% RSLogix 500 project PROGRAM_-7_BAK017.RSS, saved by version 8.30.00.16 %
PROJECT "UNTITLED"    % processor: Bul.1763 MicroLogix 1100 Series B %

PROGRAM FILES
  LAD 2 "MAIN"  4 rungs
  LAD 3 "IO"  4 rungs
  LAD 4 "SAMPL_CYCL"  2 rungs
  LAD 5 "CAL_CYCL"  14 rungs

DATA FILES
  O0 OUTPUT  4 elements
  I1 INPUT  6 elements
  S2 STATUS  66 elements
  B3 BINARY  1 elements
  T4 TIMER  3 elements
  C5 COUNTER  1 elements
  R6 CONTROL  1 elements
  N7 INTEGER  8 elements
  F8 FLOAT  7 elements

LADDER 2 "MAIN"
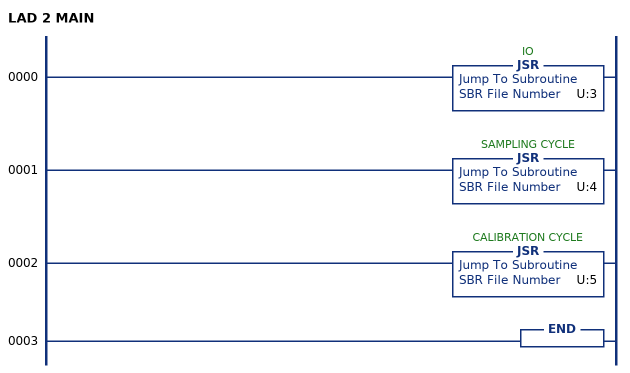
% Rung: 0 %
SOR JSR U:3 EOR
%   U:3  "IO" %
% Rung: 1 %
SOR JSR U:4 EOR
%   U:4  "SAMPLING CYCLE" %
% Rung: 2 %
SOR JSR U:5 EOR
%   U:5  "CALIBRATION CYCLE" %
% Rung: 3 %
SOR END EOR

LADDER 3 "IO"
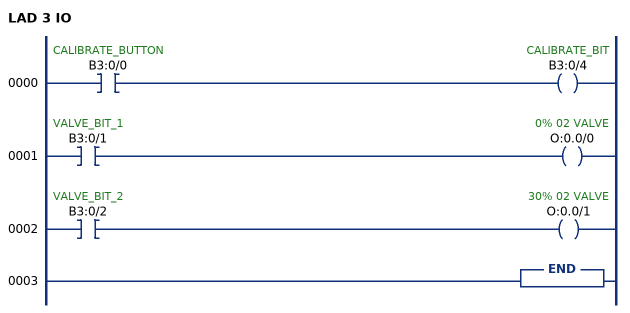
% Rung: 0 %
SOR XIC B3:0/0 OTE B3:0/4 EOR
%   B3:0/0  CALIBRATE_BUTTON %
%   B3:0/4  CALIBRATE_BIT %
% Rung: 1 %
SOR XIC B3:0/1 OTE O:0.0/0 EOR
%   B3:0/1  VALVE_BIT_1 %
%   O:0.0/0  "0% 02 VALVE" %
% Rung: 2 %
SOR XIC B3:0/2 OTE O:0.0/1 EOR
%   B3:0/2  VALVE_BIT_2 %
%   O:0.0/1  "30% 02 VALVE" %
% Rung: 3 %
SOR END EOR

LADDER 4 "SAMPL_CYCL"
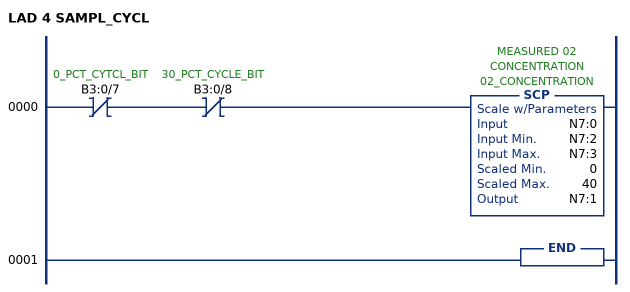
% Rung: 0 %
SOR XIO B3:0/7 XIO B3:0/8 SCP N7:0 N7:2 N7:3 0 40 N7:1 EOR
%   B3:0/7  0_PCT_CYTCL_BIT %
%   B3:0/8  30_PCT_CYCLE_BIT %
%   N7:0  02_SENSOR_VALUE  "02 SENSOR" %
%   N7:2  MIN_INPUT_0_PCT  "02 INPUT MIN 0%" %
%   N7:3  MAX_INPUT_40_PCT  "02 INPUT MAX 40%" %
%   N7:1  02_CONCENTRATION  "MEASURED 02 CONCENTRATION" %
% Rung: 1 %
SOR END EOR

LADDER 5 "CAL_CYCL"
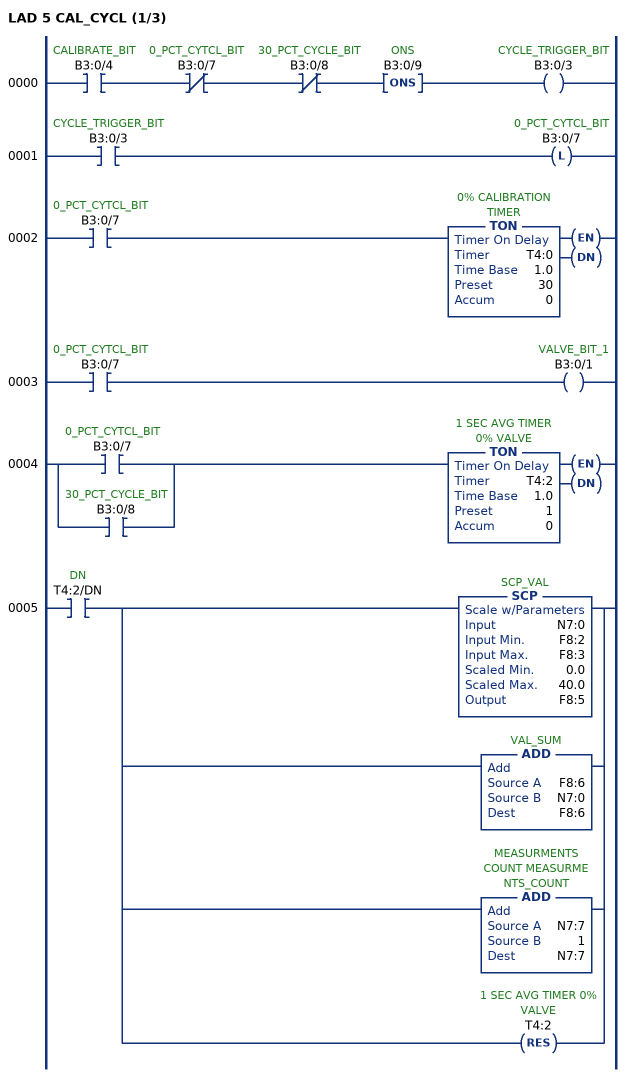
% Rung: 0 %
SOR XIC B3:0/4 XIO B3:0/7 XIO B3:0/8 ONS B3:0/9 OTE B3:0/3 EOR
%   B3:0/4  CALIBRATE_BIT %
%   B3:0/7  0_PCT_CYTCL_BIT %
%   B3:0/8  30_PCT_CYCLE_BIT %
%   B3:0/9  "ONS" %
%   B3:0/3  CYCLE_TRIGGER_BIT %
% Rung: 1 %
SOR XIC B3:0/3 OTL B3:0/7 EOR
%   B3:0/3  CYCLE_TRIGGER_BIT %
%   B3:0/7  0_PCT_CYTCL_BIT %
% Rung: 2 %
SOR XIC B3:0/7 TON T4:0 1.0 30 0 EOR
%   B3:0/7  0_PCT_CYTCL_BIT %
%   T4:0  "0% CALIBRATION TIMER" %
% Rung: 3 %
SOR XIC B3:0/7 OTE B3:0/1 EOR
%   B3:0/7  0_PCT_CYTCL_BIT %
%   B3:0/1  VALVE_BIT_1 %
% Rung: 4 %
SOR BST XIC B3:0/7 NXB XIC B3:0/8 BND TON T4:2 1.0 1 0 EOR
%   B3:0/7  0_PCT_CYTCL_BIT %
%   B3:0/8  30_PCT_CYCLE_BIT %
%   T4:2  "1 SEC AVG TIMER 0% VALVE" %
% Rung: 5 %
SOR XIC T4:2/DN BST SCP N7:0 F8:2 F8:3 0.0 40.0 F8:5 NXB ADD F8:6 N7:0 F8:6 NXB ADD N7:7 1 N7:7 NXB RES T4:2 BND EOR
%   T4:2/DN  DN %
%   N7:0  02_SENSOR_VALUE  "02 SENSOR" %
%   F8:2  INPUT_MIN %
%   F8:3  INPUT_MAX %
%   F8:5  SCP_VAL %
%   F8:6  VAL_SUM %
%   N7:7  MEASURMENTS_COUNT  "MEASURMENTS COUNT" %
%   T4:2  "1 SEC AVG TIMER 0% VALVE" %

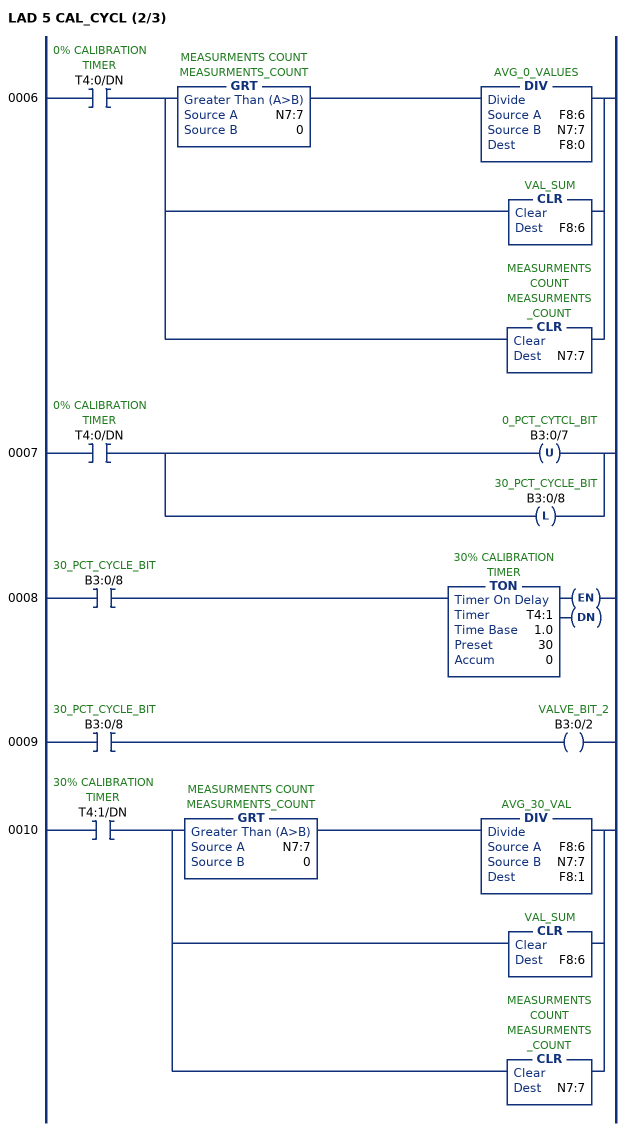
% Rung: 6 %
SOR XIC T4:0/DN BST GRT N7:7 0 DIV F8:6 N7:7 F8:0 NXB CLR F8:6 NXB CLR N7:7 BND EOR
%   T4:0/DN  "0% CALIBRATION TIMER" %
%   N7:7  MEASURMENTS_COUNT  "MEASURMENTS COUNT" %
%   F8:6  VAL_SUM %
%   F8:0  AVG_0_VALUES %
% Rung: 7 %
SOR XIC T4:0/DN BST OTU B3:0/7 NXB OTL B3:0/8 BND EOR
%   T4:0/DN  "0% CALIBRATION TIMER" %
%   B3:0/7  0_PCT_CYTCL_BIT %
%   B3:0/8  30_PCT_CYCLE_BIT %
% Rung: 8 %
SOR XIC B3:0/8 TON T4:1 1.0 30 0 EOR
%   B3:0/8  30_PCT_CYCLE_BIT %
%   T4:1  "30% CALIBRATION TIMER" %
% Rung: 9 %
SOR XIC B3:0/8 OTE B3:0/2 EOR
%   B3:0/8  30_PCT_CYCLE_BIT %
%   B3:0/2  VALVE_BIT_2 %
% Rung: 10 %
SOR XIC T4:1/DN BST GRT N7:7 0 DIV F8:6 N7:7 F8:1 NXB CLR F8:6 NXB CLR N7:7 BND EOR
%   T4:1  "30% CALIBRATION TIMER" %
%   N7:7  MEASURMENTS_COUNT  "MEASURMENTS COUNT" %
%   F8:6  VAL_SUM %
%   F8:1  AVG_30_VAL %

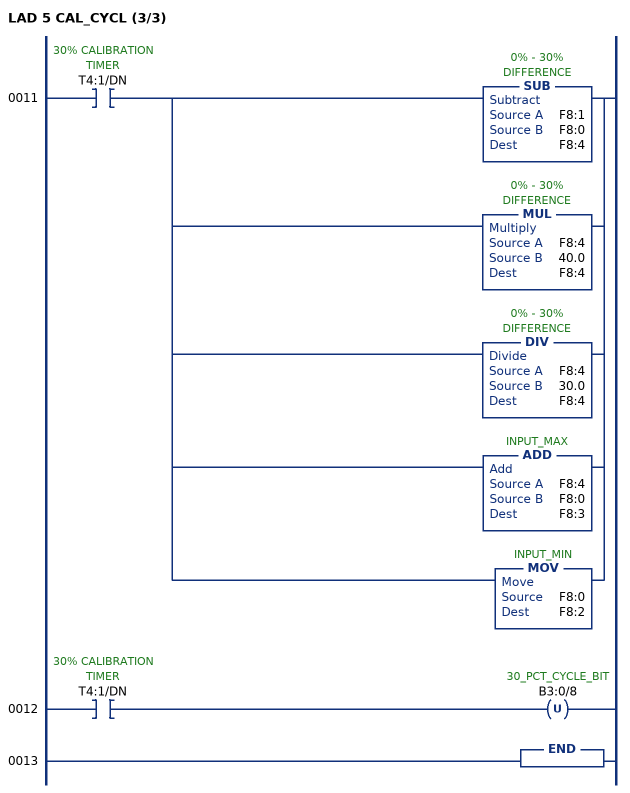
% Rung: 11 %
SOR XIC T4:1/DN BST SUB F8:1 F8:0 F8:4 NXB MUL F8:4 40.0 F8:4 NXB DIV F8:4 30.0 F8:4 NXB ADD F8:4 F8:0 F8:3 NXB MOV F8:0 F8:2 BND EOR
%   T4:1  "30% CALIBRATION TIMER" %
%   F8:1  AVG_30_VAL %
%   F8:0  AVG_0_VALUES %
%   F8:4  "0% - 30% DIFFERENCE" %
%   F8:3  INPUT_MAX %
%   F8:2  INPUT_MIN %
% Rung: 12 %
SOR XIC T4:1/DN OTU B3:0/8 EOR
%   T4:1  "30% CALIBRATION TIMER" %
%   B3:0/8  30_PCT_CYCLE_BIT %
% Rung: 13 %
SOR END EOR

OTHER DOCUMENTED ADDRESSES
  B3:0/5  "ONS"
  B3:0/6  ACTIVE_CYCLE_BIT
  F7:5  "CONCETRATION_PER_SEC"
  F7:6  "SUM OF VALUES"
  F7:8  "CYCLE_AVG"
  F7:9  MIN_AVG_VALUE
  F8:7  AVG_CYCL_VAL
  N7:5  "CONCETRATION_SECOND"

DATA TABLE (non-zero values as saved)
DATA T4
% .PRE .ACC %
% T4:0 % 30 0
% T4:1 % 30 0
% T4:2 % 1 0
DATA N7
% N7:0 % 14633 36 0 16383 0 0 0 0
DATA F8
% F8:0 % 100 11000 100 14633.33 14533.33
% F8:5 % 26.74704 0
